// TIA Portal V20 export
DATA_BLOCK "T2_Datos_Nuevos"   // DB40922
{ S7_Optimized_Access := 'TRUE' }
AUTHOR : IA
FAMILY : PRUEBA
VERSION : 0.1
// Prueba IA 2: datos de las pruebas nuevas
// stored: AutoNumber false
   VAR
      Mul_Out : Int;
      Div_Out : Int;
      Suma_Out : Int;
   END_VAR
BEGIN
END_DATA_BLOCK
